DATA_BLOCK "DB SENSOR CHECK"
TITLE =
VERSION : 0.1


  STRUCT
   B5_1 : "Sensor Check Struct";
   B5_2 : "Sensor Check Struct";
   B5_4 : "Sensor Check Struct";
   B5_5 : "Sensor Check Struct";
   B6_0 : "Sensor Check Struct";
   B6_1 : "Sensor Check Struct";
   B6_2 : "Sensor Check Struct";
   B6_4 : "Sensor Check Struct";
   B6_7 : "Sensor Check Struct";
   B7_0 : "Sensor Check Struct";
   B7_1 : "Sensor Check Struct";
   B7_2 : "Sensor Check Struct";
   B7_3 : "Sensor Check Struct";
   B7_4 : "Sensor Check Struct";
   B8_2 : "Sensor Check Struct";
   B9_6 : "Sensor Check Struct";
   B9_7 : "Sensor Check Struct";
   B10_3 : "Sensor Check Struct";
   B10_4 : "Sensor Check Struct";
   B10_5 : "Sensor Check Struct";
   B10_6 : "Sensor Check Struct";
   B10_7 : "Sensor Check Struct";
   B11_0 : "Sensor Check Struct";
   B11_1 : "Sensor Check Struct";
   B12_3 : "Sensor Check Struct";
   B13_0 : "Sensor Check Struct";
   B15_4 : "Sensor Check Struct";
   B15_5 : "Sensor Check Struct";
   B15_6 : "Sensor Check Struct";
   B15_7 : "Sensor Check Struct";
   B35_2 : "Sensor Check Struct";
   B35_3 : "Sensor Check Struct";
   B35_4 : "Sensor Check Struct";
   B11_2 : "Sensor Check Struct";
   Z2040 : BOOL ;
   M052 : BOOL ;
   M1122 : BOOL ;
   M1123 : BOOL ;
   M1124 : BOOL ;
   M1125 : BOOL ;
   M1126 : BOOL ;
   M1127 : BOOL ;
  END_STRUCT ;
BEGIN
   B5_1.Rising_Pulse_1 := FALSE;
   B5_1.Rising_Pulse_2 := FALSE;
   B5_1.Memory_Bit_1 := FALSE;
   B5_1.Memory_Bit_2 := FALSE;
   B5_1.Word_buffer := 0;
   B5_1.Word_Result := 0;
   B5_2.Rising_Pulse_1 := FALSE;
   B5_2.Rising_Pulse_2 := FALSE;
   B5_2.Memory_Bit_1 := FALSE;
   B5_2.Memory_Bit_2 := FALSE;
   B5_2.Word_buffer := 0;
   B5_2.Word_Result := 0;
   B5_4.Rising_Pulse_1 := FALSE;
   B5_4.Rising_Pulse_2 := FALSE;
   B5_4.Memory_Bit_1 := FALSE;
   B5_4.Memory_Bit_2 := FALSE;
   B5_4.Word_buffer := 0;
   B5_4.Word_Result := 0;
   B5_5.Rising_Pulse_1 := FALSE;
   B5_5.Rising_Pulse_2 := FALSE;
   B5_5.Memory_Bit_1 := FALSE;
   B5_5.Memory_Bit_2 := FALSE;
   B5_5.Word_buffer := 0;
   B5_5.Word_Result := 0;
   B6_0.Rising_Pulse_1 := FALSE;
   B6_0.Rising_Pulse_2 := FALSE;
   B6_0.Memory_Bit_1 := FALSE;
   B6_0.Memory_Bit_2 := FALSE;
   B6_0.Word_buffer := 0;
   B6_0.Word_Result := 0;
   B6_1.Rising_Pulse_1 := FALSE;
   B6_1.Rising_Pulse_2 := FALSE;
   B6_1.Memory_Bit_1 := FALSE;
   B6_1.Memory_Bit_2 := FALSE;
   B6_1.Word_buffer := 0;
   B6_1.Word_Result := 0;
   B6_2.Rising_Pulse_1 := FALSE;
   B6_2.Rising_Pulse_2 := FALSE;
   B6_2.Memory_Bit_1 := FALSE;
   B6_2.Memory_Bit_2 := FALSE;
   B6_2.Word_buffer := 0;
   B6_2.Word_Result := 0;
   B6_4.Rising_Pulse_1 := FALSE;
   B6_4.Rising_Pulse_2 := FALSE;
   B6_4.Memory_Bit_1 := FALSE;
   B6_4.Memory_Bit_2 := FALSE;
   B6_4.Word_buffer := 0;
   B6_4.Word_Result := 0;
   B6_7.Rising_Pulse_1 := FALSE;
   B6_7.Rising_Pulse_2 := FALSE;
   B6_7.Memory_Bit_1 := FALSE;
   B6_7.Memory_Bit_2 := FALSE;
   B6_7.Word_buffer := 0;
   B6_7.Word_Result := 0;
   B7_0.Rising_Pulse_1 := FALSE;
   B7_0.Rising_Pulse_2 := FALSE;
   B7_0.Memory_Bit_1 := FALSE;
   B7_0.Memory_Bit_2 := FALSE;
   B7_0.Word_buffer := 0;
   B7_0.Word_Result := 0;
   B7_1.Rising_Pulse_1 := FALSE;
   B7_1.Rising_Pulse_2 := FALSE;
   B7_1.Memory_Bit_1 := FALSE;
   B7_1.Memory_Bit_2 := FALSE;
   B7_1.Word_buffer := 0;
   B7_1.Word_Result := 0;
   B7_2.Rising_Pulse_1 := FALSE;
   B7_2.Rising_Pulse_2 := FALSE;
   B7_2.Memory_Bit_1 := FALSE;
   B7_2.Memory_Bit_2 := FALSE;
   B7_2.Word_buffer := 0;
   B7_2.Word_Result := 0;
   B7_3.Rising_Pulse_1 := FALSE;
   B7_3.Rising_Pulse_2 := FALSE;
   B7_3.Memory_Bit_1 := FALSE;
   B7_3.Memory_Bit_2 := FALSE;
   B7_3.Word_buffer := 0;
   B7_3.Word_Result := 0;
   B7_4.Rising_Pulse_1 := FALSE;
   B7_4.Rising_Pulse_2 := FALSE;
   B7_4.Memory_Bit_1 := FALSE;
   B7_4.Memory_Bit_2 := FALSE;
   B7_4.Word_buffer := 0;
   B7_4.Word_Result := 0;
   B8_2.Rising_Pulse_1 := FALSE;
   B8_2.Rising_Pulse_2 := FALSE;
   B8_2.Memory_Bit_1 := FALSE;
   B8_2.Memory_Bit_2 := FALSE;
   B8_2.Word_buffer := 0;
   B8_2.Word_Result := 0;
   B9_6.Rising_Pulse_1 := FALSE;
   B9_6.Rising_Pulse_2 := FALSE;
   B9_6.Memory_Bit_1 := FALSE;
   B9_6.Memory_Bit_2 := FALSE;
   B9_6.Word_buffer := 0;
   B9_6.Word_Result := 0;
   B9_7.Rising_Pulse_1 := FALSE;
   B9_7.Rising_Pulse_2 := FALSE;
   B9_7.Memory_Bit_1 := FALSE;
   B9_7.Memory_Bit_2 := FALSE;
   B9_7.Word_buffer := 0;
   B9_7.Word_Result := 0;
   B10_3.Rising_Pulse_1 := FALSE;
   B10_3.Rising_Pulse_2 := FALSE;
   B10_3.Memory_Bit_1 := FALSE;
   B10_3.Memory_Bit_2 := FALSE;
   B10_3.Word_buffer := 0;
   B10_3.Word_Result := 0;
   B10_4.Rising_Pulse_1 := FALSE;
   B10_4.Rising_Pulse_2 := FALSE;
   B10_4.Memory_Bit_1 := FALSE;
   B10_4.Memory_Bit_2 := FALSE;
   B10_4.Word_buffer := 0;
   B10_4.Word_Result := 0;
   B10_5.Rising_Pulse_1 := FALSE;
   B10_5.Rising_Pulse_2 := FALSE;
   B10_5.Memory_Bit_1 := FALSE;
   B10_5.Memory_Bit_2 := FALSE;
   B10_5.Word_buffer := 0;
   B10_5.Word_Result := 0;
   B10_6.Rising_Pulse_1 := FALSE;
   B10_6.Rising_Pulse_2 := FALSE;
   B10_6.Memory_Bit_1 := FALSE;
   B10_6.Memory_Bit_2 := FALSE;
   B10_6.Word_buffer := 0;
   B10_6.Word_Result := 0;
   B10_7.Rising_Pulse_1 := FALSE;
   B10_7.Rising_Pulse_2 := FALSE;
   B10_7.Memory_Bit_1 := FALSE;
   B10_7.Memory_Bit_2 := FALSE;
   B10_7.Word_buffer := 0;
   B10_7.Word_Result := 0;
   B11_0.Rising_Pulse_1 := FALSE;
   B11_0.Rising_Pulse_2 := FALSE;
   B11_0.Memory_Bit_1 := FALSE;
   B11_0.Memory_Bit_2 := FALSE;
   B11_0.Word_buffer := 0;
   B11_0.Word_Result := 0;
   B11_1.Rising_Pulse_1 := FALSE;
   B11_1.Rising_Pulse_2 := FALSE;
   B11_1.Memory_Bit_1 := FALSE;
   B11_1.Memory_Bit_2 := FALSE;
   B11_1.Word_buffer := 0;
   B11_1.Word_Result := 0;
   B12_3.Rising_Pulse_1 := FALSE;
   B12_3.Rising_Pulse_2 := FALSE;
   B12_3.Memory_Bit_1 := FALSE;
   B12_3.Memory_Bit_2 := FALSE;
   B12_3.Word_buffer := 0;
   B12_3.Word_Result := 0;
   B13_0.Rising_Pulse_1 := FALSE;
   B13_0.Rising_Pulse_2 := FALSE;
   B13_0.Memory_Bit_1 := FALSE;
   B13_0.Memory_Bit_2 := FALSE;
   B13_0.Word_buffer := 0;
   B13_0.Word_Result := 0;
   B15_4.Rising_Pulse_1 := FALSE;
   B15_4.Rising_Pulse_2 := FALSE;
   B15_4.Memory_Bit_1 := FALSE;
   B15_4.Memory_Bit_2 := FALSE;
   B15_4.Word_buffer := 0;
   B15_4.Word_Result := 0;
   B15_5.Rising_Pulse_1 := FALSE;
   B15_5.Rising_Pulse_2 := FALSE;
   B15_5.Memory_Bit_1 := FALSE;
   B15_5.Memory_Bit_2 := FALSE;
   B15_5.Word_buffer := 0;
   B15_5.Word_Result := 0;
   B15_6.Rising_Pulse_1 := FALSE;
   B15_6.Rising_Pulse_2 := FALSE;
   B15_6.Memory_Bit_1 := FALSE;
   B15_6.Memory_Bit_2 := FALSE;
   B15_6.Word_buffer := 0;
   B15_6.Word_Result := 0;
   B15_7.Rising_Pulse_1 := FALSE;
   B15_7.Rising_Pulse_2 := FALSE;
   B15_7.Memory_Bit_1 := FALSE;
   B15_7.Memory_Bit_2 := FALSE;
   B15_7.Word_buffer := 0;
   B15_7.Word_Result := 0;
   B35_2.Rising_Pulse_1 := FALSE;
   B35_2.Rising_Pulse_2 := FALSE;
   B35_2.Memory_Bit_1 := FALSE;
   B35_2.Memory_Bit_2 := FALSE;
   B35_2.Word_buffer := 0;
   B35_2.Word_Result := 0;
   B35_3.Rising_Pulse_1 := FALSE;
   B35_3.Rising_Pulse_2 := FALSE;
   B35_3.Memory_Bit_1 := FALSE;
   B35_3.Memory_Bit_2 := FALSE;
   B35_3.Word_buffer := 0;
   B35_3.Word_Result := 0;
   B35_4.Rising_Pulse_1 := FALSE;
   B35_4.Rising_Pulse_2 := FALSE;
   B35_4.Memory_Bit_1 := FALSE;
   B35_4.Memory_Bit_2 := FALSE;
   B35_4.Word_buffer := 0;
   B35_4.Word_Result := 0;
   B11_2.Rising_Pulse_1 := FALSE;
   B11_2.Rising_Pulse_2 := FALSE;
   B11_2.Memory_Bit_1 := FALSE;
   B11_2.Memory_Bit_2 := FALSE;
   B11_2.Word_buffer := 0;
   B11_2.Word_Result := 0;
   Z2040 := FALSE;
   M052 := FALSE;
   M1122 := FALSE;
   M1123 := FALSE;
   M1124 := FALSE;
   M1125 := FALSE;
   M1126 := FALSE;
   M1127 := FALSE;
END_DATA_BLOCK
